// TIA Portal V20 export
// export: Created 2026-10-12T05:06:09.0081338Z, ExportSetting WithDefaults, DisplayName Totally Integrated Automation Portal, DisplayVersion V20, DisplayName TIA Portal Openness, DisplayVersion V20, DisplayName TIA Portal Teamcenter Gateway, DisplayVersion V20, DisplayName TIA Portal Version Control Interface, DisplayVersion V20, DisplayName SINAMICS Startdrive Advanced, DisplayVersion V20 SP1 Update 2, DisplayName SINAMICS Startdrive G110M, G120, G120C, G120D, G120P, G115D, DisplayVersion V20 SP1 Update 2, DisplayName SINAMICS Startdrive G130, G150, S120, S150, SINAMICS MV, G220, S200, S210, DisplayVersion V20 SP1 Update 2, DisplayName STEP 7 Professional, DisplayVersion V20, DisplayName STEP 7 Safety, DisplayVersion V20, DisplayName WinCC Basic/Comfort/Advanced, DisplayVersion V20, DisplayName WinCC Professional, DisplayVersion V20, DisplayName WinCC Unified, DisplayVersion V20
TYPE "ST_ConfigSetInfo"
// stored: IsFailsafeCompliant false
   STRUCT
      Used : Bool;
      SetName : String[80];
      RootIdentity : String[80];
      SetSchema : UInt;
      ConfigRev : UDInt;
      Kind : DInt;
      ModelCode : String[64];
      RecordCount : Int;
      CreatedAt : LDT;
      TimeSynchronized : Bool;
   END_STRUCT;
END_TYPE
